(* IEC 61131-3 sources: STEPROBOT/docs/auto_job_r6_4/plc, 18 files *)

(* ---- GVL_FileBridge.st ---- *)
{attribute 'qualified_only'}
VAR_GLOBAL PERSISTENT RETAIN
    (* Reserve these MW ranges in the FIELD project before importing. *)
    aCommand AT %MW6000 : ARRAY[0..119] OF WORD;
    aHeartbeat AT %MW6120 : ARRAY[0..4] OF WORD;
    aStatus AT %MW6200 : ARRAY[0..63] OF WORD;
END_VAR
VAR_GLOBAL
    (* LOCAL configuration only. Never map credentials/permit to Modbus. *)
    xFileTransferPermit : BOOL := FALSE;
    xReset : BOOL := FALSE;
    sFtpUser : STRING(64) := '';
    sFtpPassword : STRING(64) := '';
    aBuffer : ARRAY[0..1048575] OF BYTE;
    (* One-time LOCAL commissioning: exact existing project already bound to these manual service and one auto GDI number.
       This mode reuses bindings. It never edits robot system configuration. *)
    xFixedMappingConfirmed : BOOL := FALSE;
    sFixedProject : STRING(64) := 'pcjob_manual_r63.sr';
    uiFixedCapture : UINT := UINT#10;
    uiFixedPath : UINT := UINT#11;
    uiAutoCapacity : UINT := UINT#15;
    (* Nonretained: a reboot or failed update never authorizes a partly updated project. *)
    xFixedUpdateBusy : BOOL;
    xFixedReady : BOOL;
    xFixedIdle : BOOL;
    aAutoTag : ARRAY[0..2] OF WORD;
END_VAR

(* ---- GVL_FileBridgeRetain.st ---- *)
{attribute 'qualified_only'}
VAR_GLOBAL PERSISTENT RETAIN
    udiBootCounter : UDINT := UDINT#0;
END_VAR

(* ---- GVL_ManualBridge.st ---- *)
{attribute 'qualified_only'}
VAR_GLOBAL PERSISTENT RETAIN
    // PC extension: no overlap with HR200..215, HR300..363 or FTP HR6000+.
    aCommand AT %MW220 : ARRAY[0..15] OF WORD;
    aStatus AT %MW400 : ARRAY[0..31] OF WORD;
END_VAR
VAR_GLOBAL
    // Local configuration. Assign ONE unused GDI slot to manual_service before setting TRUE.
    xInstalled : BOOL := FALSE;
    xServiceBindingConfirmed : BOOL := FALSE;
    uiServiceProgram : UINT := 10;
    // PRG_ManualBridge is the only writer. PRG_RobotBridge reads these requests.
    xActive : BOOL;
    xStartRequest : BOOL;
    xStopRequest : BOOL;
END_VAR

(* ---- GVL_ParamProbe.st ---- *)
{attribute 'qualified_only'}
VAR_GLOBAL
    // Mapped to existing ParamProbe_Write FC16 offset4 length4. Single writer: PRG_ManualBridge.
    aParamTx : ARRAY[0..3] OF WORD;
END_VAR

(* ---- GVL_RobotBridge.st ---- *)
{attribute 'qualified_only'}
VAR_GLOBAL PERSISTENT RETAIN
    // PC <-> PLC. Inovance native Modbus TCP slave: MWn <-> HR offset n.
    // Commission by reading HR300=16#4D42 and HR301=2 before permitting motion.
    aHostCmd AT %MW200 : ARRAY[0..15] OF WORD;
    aHostStatus AT %MW300 : ARRAY[0..63] OF WORD;

END_VAR

VAR_GLOBAL
    // PLC master -> STEP slave: FC04 / offset 0 / 32 WORD.
    aRobotRx : ARRAY[0..31] OF WORD;
    // PLC master -> STEP slave: ONE FC16 / offset 0 / 2 WORDs.
    // Map BOTH aRobotTx[0] and aRobotTx[1], NOT wRobotTxControl alone.
    aRobotTx : ARRAY[0..1] OF WORD;
    wRobotTxControl : WORD; // first-word diagnostic alias, not a separate channel

    // Local commissioning/operation inputs. Do not map these into aHostCmd.
    xCommissioned : BOOL := FALSE;
    // Set locally ONLY after checking DI49..56 and the GDI program bindings.
    xGdiProgramMappingConfirmed : BOOL := FALSE;
    xRemotePermit : BOOL := FALSE;
    // Optional native master/channel fault. FALSE leaves DO42 watchdog in use.
    xNativeModbusError : BOOL := FALSE;

    // Published live diagnostics.
    xRobotLinkOK : BOOL;
    xRobotRunning : BOOL;
    xRobotPaused : BOOL;
    xRobotStopped : BOOL;
    xRobotEnabled : BOOL;
    xRobotAlarm : BOOL;
    xRobotEmergency : BOOL;
    xRobotExternalAuto : BOOL;
    xHostRegistered : BOOL;
    xHostAlive : BOOL;
    xBusy : BOOL;
    xStopInterlock : BOOL;
    xLoadOperatorConfirmed : BOOL;
    uiFixedJobGuardVersion : UINT;
END_VAR

(* ---- GVL_RobotBridgeRetain.st ---- *)
{attribute 'qualified_only'}
VAR_GLOBAL PERSISTENT RETAIN
    // Incremented on application initialization, not on every scan.
    // Also require a fresh registration; a cold reset can reset RETAIN memory.
    udiBootCounter : UDINT := 0;
END_VAR

(* ---- GVL_RobotJoints.st ---- *)
{attribute 'qualified_only'}
VAR_GLOBAL PERSISTENT RETAIN
    // PC reads HR500..539. Reserve this unused range in the field project.
    // The publisher rebuilds all validity metadata; retained values never grant validity.
    aStatus AT %MW500 : ARRAY[0..39] OF WORD;
END_VAR
VAR_GLOBAL
    xEnable : BOOL := TRUE;
    sRobotAddress : STRING(15) := '192.168.3.188';
    uiRobotPort : UINT := UINT#502;
    byRobotUnit : BYTE := BYTE#1;
    // Local commissioning only: compare all six axes with the pendant.
    // FALSE = first register is the low half of IEEE754 REAL.
    xHighWordFirst : BOOL := FALSE;
END_VAR

(* ---- F_AutoFileIndex.st ---- *)
FUNCTION F_AutoFileIndex : UINT
VAR_INPUT
    sName : STRING(64);
END_VAR
F_AutoFileIndex := UINT#0;
IF sName = 'auto_main.srd' THEN F_AutoFileIndex := UINT#1; END_IF;
IF sName = 'auto_main.srp' THEN F_AutoFileIndex := UINT#2; END_IF;
IF sName = 'auto_01.srd' THEN F_AutoFileIndex := UINT#3; END_IF;
IF sName = 'auto_01.srp' THEN F_AutoFileIndex := UINT#4; END_IF;
IF sName = 'auto_02.srd' THEN F_AutoFileIndex := UINT#5; END_IF;
IF sName = 'auto_02.srp' THEN F_AutoFileIndex := UINT#6; END_IF;
IF sName = 'auto_03.srd' THEN F_AutoFileIndex := UINT#7; END_IF;
IF sName = 'auto_03.srp' THEN F_AutoFileIndex := UINT#8; END_IF;
IF sName = 'auto_04.srd' THEN F_AutoFileIndex := UINT#9; END_IF;
IF sName = 'auto_04.srp' THEN F_AutoFileIndex := UINT#10; END_IF;
IF sName = 'auto_05.srd' THEN F_AutoFileIndex := UINT#11; END_IF;
IF sName = 'auto_05.srp' THEN F_AutoFileIndex := UINT#12; END_IF;
IF sName = 'auto_06.srd' THEN F_AutoFileIndex := UINT#13; END_IF;
IF sName = 'auto_06.srp' THEN F_AutoFileIndex := UINT#14; END_IF;
IF sName = 'auto_07.srd' THEN F_AutoFileIndex := UINT#15; END_IF;
IF sName = 'auto_07.srp' THEN F_AutoFileIndex := UINT#16; END_IF;
IF sName = 'auto_08.srd' THEN F_AutoFileIndex := UINT#17; END_IF;
IF sName = 'auto_08.srp' THEN F_AutoFileIndex := UINT#18; END_IF;
IF sName = 'auto_09.srd' THEN F_AutoFileIndex := UINT#19; END_IF;
IF sName = 'auto_09.srp' THEN F_AutoFileIndex := UINT#20; END_IF;
IF sName = 'auto_10.srd' THEN F_AutoFileIndex := UINT#21; END_IF;
IF sName = 'auto_10.srp' THEN F_AutoFileIndex := UINT#22; END_IF;
IF sName = 'auto_11.srd' THEN F_AutoFileIndex := UINT#23; END_IF;
IF sName = 'auto_11.srp' THEN F_AutoFileIndex := UINT#24; END_IF;
IF sName = 'auto_12.srd' THEN F_AutoFileIndex := UINT#25; END_IF;
IF sName = 'auto_12.srp' THEN F_AutoFileIndex := UINT#26; END_IF;
IF sName = 'auto_13.srd' THEN F_AutoFileIndex := UINT#27; END_IF;
IF sName = 'auto_13.srp' THEN F_AutoFileIndex := UINT#28; END_IF;
IF sName = 'auto_14.srd' THEN F_AutoFileIndex := UINT#29; END_IF;
IF sName = 'auto_14.srp' THEN F_AutoFileIndex := UINT#30; END_IF;
IF sName = 'auto_15.srd' THEN F_AutoFileIndex := UINT#31; END_IF;
IF sName = 'auto_15.srp' THEN F_AutoFileIndex := UINT#32; END_IF;
END_FUNCTION

(* ---- F_FileCrc32.st ---- *)
FUNCTION F_FileCrc32 : UDINT
VAR_INPUT
    pData : POINTER TO BYTE;
    uiCount : UINT;
    udiSeed : UDINT;
END_VAR
VAR
    udiCrc : UDINT;
    uiI : UINT;
    uiBit : UINT;
END_VAR
(* Running reflected CRC-32. Caller supplies initial FFFFFFFF and final XOR. *)
udiCrc := udiSeed;
IF uiCount > UINT#0 THEN
    FOR uiI := UINT#0 TO uiCount - UINT#1 DO
        udiCrc := udiCrc XOR BYTE_TO_UDINT(pData[uiI]);
        FOR uiBit := UINT#0 TO UINT#7 DO
            IF (udiCrc AND UDINT#1) <> UDINT#0 THEN
                udiCrc := SHR(udiCrc, 1) XOR UDINT#16#EDB88320;
            ELSE
                udiCrc := SHR(udiCrc, 1);
            END_IF;
        END_FOR;
    END_FOR;
END_IF;
F_FileCrc32 := udiCrc;
END_FUNCTION

(* ---- F_FileCrc32Fast.st ---- *)
FUNCTION F_FileCrc32Fast : UDINT
VAR_INPUT
    pData : POINTER TO BYTE;
    uiCount : UINT;
    udiSeed : UDINT;
END_VAR
VAR
    udiCrc : UDINT;
    udiTable : UDINT;
    uiI : UINT;
    uiNibble : UINT;
END_VAR
(* Reflected CRC32, two nibble lookups per byte; no initialization scan. *)
udiCrc := udiSeed;
IF uiCount > UINT#0 THEN
    FOR uiI := UINT#0 TO uiCount - UINT#1 DO
        udiCrc := udiCrc XOR BYTE_TO_UDINT(pData[uiI]);
        FOR uiNibble := UINT#0 TO UINT#1 DO
            CASE udiCrc AND UDINT#15 OF
                0: udiTable := UDINT#16#00000000;
                1: udiTable := UDINT#16#1DB71064;
                2: udiTable := UDINT#16#3B6E20C8;
                3: udiTable := UDINT#16#26D930AC;
                4: udiTable := UDINT#16#76DC4190;
                5: udiTable := UDINT#16#6B6B51F4;
                6: udiTable := UDINT#16#4DB26158;
                7: udiTable := UDINT#16#5005713C;
                8: udiTable := UDINT#16#EDB88320;
                9: udiTable := UDINT#16#F00F9344;
                10: udiTable := UDINT#16#D6D6A3E8;
                11: udiTable := UDINT#16#CB61B38C;
                12: udiTable := UDINT#16#9B64C2B0;
                13: udiTable := UDINT#16#86D3D2D4;
                14: udiTable := UDINT#16#A00AE278;
                15: udiTable := UDINT#16#BDBDF21C;
            END_CASE;
            udiCrc := SHR(udiCrc, 4) XOR udiTable;
        END_FOR;
    END_FOR;
END_IF;
F_FileCrc32Fast := udiCrc;
END_FUNCTION

(* ---- F_FileNameValid.st ---- *)
FUNCTION F_FileNameValid : BOOL
VAR_INPUT
    sName : STRING(64);
    xProject : BOOL;
END_VAR
VAR
    pName : POINTER TO BYTE;
    uiI : UINT;
    uiBaseLength : UINT;
    xValid : BOOL;
    xChar : BOOL;
END_VAR
(* Flat lowercase ASCII names; no slash, CR/LF, spaces, or extra dots. *)
xValid := FALSE;
uiBaseLength := UINT#0;
IF xProject THEN
    IF (LEFT(sName, 6) = 'pcjob_') AND (RIGHT(sName, 3) = '.sr')
        AND (LEN(sName) >= 12) AND (LEN(sName) <= 48) THEN
        uiBaseLength := INT_TO_UINT(LEN(sName)) - UINT#3;
    END_IF;
ELSE
    IF (LEN(sName) >= 5) AND (LEN(sName) <= 48) THEN
        IF (RIGHT(sName, 4) = '.srp') OR (RIGHT(sName, 4) = '.srd')
            OR (RIGHT(sName, 4) = '.txt') THEN
            uiBaseLength := INT_TO_UINT(LEN(sName)) - UINT#4;
        END_IF;
    END_IF;
END_IF;
IF uiBaseLength > UINT#0 THEN
    xValid := TRUE;
    pName := ADR(sName);
    FOR uiI := UINT#0 TO uiBaseLength - UINT#1 DO
        xChar := ((pName[uiI] >= BYTE#97) AND (pName[uiI] <= BYTE#122))
            OR ((pName[uiI] >= BYTE#48) AND (pName[uiI] <= BYTE#57))
            OR (pName[uiI] = BYTE#95);
        IF NOT xChar THEN xValid := FALSE; END_IF;
    END_FOR;
END_IF;
F_FileNameValid := xValid;
END_FUNCTION

(* ---- F_FixedFileValid.st ---- *)
FUNCTION F_FixedFileValid : BOOL
VAR_INPUT
    sName : STRING(64);
END_VAR
F_FixedFileValid := F_AutoFileIndex(sName) > UINT#0;
END_FUNCTION

(* ---- FB_FileFtp.st ---- *)
FUNCTION_BLOCK FB_FileFtp
VAR_INPUT
    xStart : BOOL;
    xAbort : BOOL;
    pBuffer : POINTER TO BYTE;
    udiSize : UDINT;
    sProject : STRING(64);
    sFile : STRING(64);
    xCreateProject : BOOL;
    xReplaceFixed : BOOL;
    xVerifyOnly : BOOL;
    udiVerifyCrc : UDINT;
    sUser : STRING(64);
    sPassword : STRING(64);
END_VAR
VAR CONSTANT
    cdiControlID : DINT := DINT#245;
    cdiDataID : DINT := DINT#246;
END_VAR
VAR_OUTPUT
    xDone : BOOL := FALSE;
    xTestPassed : BOOL := FALSE;
    xError : BOOL := FALSE;
    xLoginOk : BOOL := FALSE;
    xBaseDirOk : BOOL := FALSE;
    xScratchCreated : BOOL := FALSE;
    xUploadComplete : BOOL := FALSE;
    xReadbackComplete : BOOL := FALSE;
    xContentMatch : BOOL := FALSE;
    xQuitOk : BOOL := FALSE;
    xCleanupOk : BOOL := FALSE;
    uiStep : UINT := UINT#0;
    uiErrorStage : UINT := UINT#0;
    wErrorID : WORD := WORD#0;
    wDataCloseErrorID : WORD := WORD#0;
    wControlCloseErrorID : WORD := WORD#0;
    udiExpectedBytes : UDINT := UDINT#0;
    udiUploadedBytes : UDINT := UDINT#0;
    udiReadbackBytes : UDINT := UDINT#0;
    uiReplyCode : UINT := UINT#0;
    uiUserReplyCode : UINT := UINT#0;
    uiPassReplyCode : UINT := UINT#0;
    uiBaseDirReplyCode : UINT := UINT#0;
    uiNameCheckReplyCode : UINT := UINT#0;
    uiMkdReplyCode : UINT := UINT#0;
    uiStorReplyCode : UINT := UINT#0;
    uiUploadCompleteCode : UINT := UINT#0;
    uiRetrReplyCode : UINT := UINT#0;
    uiDownloadCompleteCode : UINT := UINT#0;
    uiPasvPort : UINT := UINT#0;
    wReadbackEndStatus : WORD := WORD#0;
    sRemotePath : STRING(160);
    sLastReply : STRING(255);
    sMkdReply : STRING(255);
    sPasvReply : STRING(255);
    sUploadReply : STRING(255);
    sDownloadReply : STRING(255);
    xControlOwned : BOOL := FALSE;
    xDataOwned : BOOL := FALSE;
    xUploadDataConnected : BOOL := FALSE;
    xDownloadDataConnected : BOOL := FALSE;
    xLineTruncated : BOOL := FALSE;

END_VAR
VAR
    (* Caller owns immutable buffer until xDone and clean socket closure. *)
    xAbortLatched : BOOL;
    xProgress : BOOL;
    xDirectoryReady : BOOL;
    xReplaceRun : BOOL;
    sFileRun : STRING(64);
    pBufferRun : POINTER TO BYTE;

    stControlServer : CmpHCTCPIP.ADDRESS := (strIPAddr := '192.168.3.188', uiPort := UINT#21);
    stDataServer : CmpHCTCPIP.ADDRESS;
    fbControlClient : CmpHCTCPIP.SktTCPClient;
    fbControlClose : CmpHCTCPIP.SktClose;
    fbDataClient : CmpHCTCPIP.SktTCPClient;
    fbDataClose : CmpHCTCPIP.SktClose;
    fbReplyTimeout : TON;
    fbCommandTimeout : TON;
    fbUploadTimeout : TON;
    fbReadbackTimeout : TON;
    fbDataCloseTimeout : TON;
    fbControlCloseTimeout : TON;

    xStartOld : BOOL := FALSE;
    xFail : BOOL := FALSE;
    xFinishedNow : BOOL := FALSE;
    wPendingError : WORD := WORD#0;
    uiPendingStage : UINT := UINT#0;
    uiPhase : UINT := UINT#0;
    uiNextCommand : UINT := UINT#0;
    uiTransferMode : UINT := UINT#0;
    xReplyReady : BOOL := FALSE;
    xReplyAccepted : BOOL := FALSE;
    xDigits : BOOL := FALSE;
    xMultiline : BOOL := FALSE;
    sMultilineCode : STRING(3);
    sLine : STRING(255);
    pLine : POINTER TO BYTE;
    uiLineLength : UINT := UINT#0;
    fbControlIo : FB_FileSocketIo;
    fbDataIo : FB_FileSocketIo;
    uiControlRxIndex : UINT;
    uiControlRxCount : UINT;
    uiParse : UINT;
    byControl : BYTE;
    pSendNow : POINTER TO BYTE;
    uiSendNow : UINT;
    xVerifyRun : BOOL;
    udiVerifyCrcRun : UDINT;
    udiReadbackCrc : UDINT;
    sCommand : STRING(160);
    pCommand : POINTER TO BYTE;
    uiCommandIndex : UINT := UINT#0;
    uiCommandLength : UINT := UINT#0;
    sUserRun : STRING(64);
    sPasswordRun : STRING(64);
    sScratchRun : STRING(64);
    pCredential : POINTER TO BYTE;
    uiI : UINT := UINT#0;
    xNameCharacter : BOOL := FALSE;
    xBytesMatch : BOOL := FALSE;
    xReadbackEndCandidate : BOOL := FALSE;
    xDataCloseFailed : BOOL := FALSE;
    pReply : POINTER TO BYTE;
    aPasv : ARRAY[0..5] OF UINT;
    uiPasvField : UINT := UINT#0;
    uiPasvValue : UINT := UINT#0;
    xPasvValid : BOOL := FALSE;
    xPasvInTuple : BOOL := FALSE;
    xPasvClosed : BOOL := FALSE;
    xPasvHasDigit : BOOL := FALSE;
END_VAR
(* Derived from field-passed PRG_FtpUploadProbe. New bridge is NOT field validated. *)
(* IDs 245/246 must be free; default cabinet 192.168.3.188:21. *)
(* Bounded 8192-byte I/O, exact offsets and explicit EOF. No motion commands. *)
pLine := ADR(sLine);
pCommand := ADR(sCommand);
xFail := FALSE;
xFinishedNow := FALSE;
xReplyReady := FALSE;
wPendingError := WORD#0;
uiPendingStage := UINT#20 + uiPhase * UINT#10;

pSendNow := pCommand;
uiSendNow := UINT#0;
IF uiStep = UINT#40 THEN
    pSendNow := pCommand + uiCommandIndex;
    uiSendNow := uiCommandLength - uiCommandIndex;
END_IF;
fbControlClient(xExecute := uiStep = UINT#10, diConnectID := cdiControlID,
    stServerAddress := stControlServer);
fbControlIo(xSend := uiStep = UINT#40,
    xReceive := (uiStep = UINT#20) AND (uiControlRxIndex >= uiControlRxCount),
    diConnectID := cdiControlID, pSend := pSendNow, uiSendSize := uiSendNow);
IF fbControlIo.uiCount > UINT#0 THEN
    uiControlRxIndex := UINT#0;
    uiControlRxCount := fbControlIo.uiCount;
END_IF;
pSendNow := pBufferRun;
uiSendNow := UINT#0;
IF (uiStep = UINT#60) AND (udiUploadedBytes < udiExpectedBytes) THEN
    pSendNow := pBufferRun + udiUploadedBytes;
    IF udiExpectedBytes - udiUploadedBytes > UDINT#8192 THEN
        uiSendNow := UINT#8192;
    ELSE
        uiSendNow := UDINT_TO_UINT(udiExpectedBytes - udiUploadedBytes);
    END_IF;
END_IF;
fbDataClient(xExecute := uiStep = UINT#50, diConnectID := cdiDataID,
    stServerAddress := stDataServer);
fbDataIo(xSend := (uiStep = UINT#60) AND (uiSendNow > UINT#0),
    xReceive := uiStep = UINT#70, diConnectID := cdiDataID,
    pSend := pSendNow, uiSendSize := uiSendNow);
fbDataClose(xExecute := ((uiStep = UINT#80) OR (uiStep = UINT#90))
    AND xDataOwned AND NOT xDataCloseFailed, diConnectID := cdiDataID);
fbControlClose(xExecute := (uiStep = UINT#95) AND xControlOwned,
    diConnectID := cdiControlID);
fbReplyTimeout(IN := uiStep = UINT#20, PT := T#20s);
fbCommandTimeout(IN := (uiStep = UINT#40) OR (uiStep = UINT#45), PT := T#30s);
xProgress := ((uiStep = UINT#60) AND (fbDataIo.uiSent > UINT#0))
    OR ((uiStep = UINT#70) AND (fbDataIo.uiCount > UINT#0));
fbUploadTimeout(IN := ((uiStep = UINT#60) OR (uiStep = UINT#65)) AND NOT xProgress,
    PT := T#30s);
fbReadbackTimeout(IN := (uiStep = UINT#70) AND NOT xProgress, PT := T#30s);
fbDataCloseTimeout(IN := ((uiStep = UINT#80) OR (uiStep = UINT#90))
    AND xDataOwned AND NOT xDataCloseFailed, PT := T#5s);
fbControlCloseTimeout(IN := uiStep = UINT#95, PT := T#5s);

(* Bounded control-reply parser; identical-code SPACE terminates multiline replies. *)
IF (uiStep = UINT#20) AND NOT fbControlIo.xError THEN
    IF uiControlRxIndex < uiControlRxCount THEN
    FOR uiParse := uiControlRxIndex TO uiControlRxCount - UINT#1 DO
      IF (uiControlRxIndex < uiControlRxCount) AND NOT xReplyReady AND NOT xFail THEN
        byControl := fbControlIo.aRecv[uiControlRxIndex];
        uiControlRxIndex := uiControlRxIndex + UINT#1;
        IF byControl = BYTE#10 THEN
            IF uiLineLength > UINT#0 THEN
                IF pLine[uiLineLength - UINT#1] = BYTE#13 THEN
                    uiLineLength := uiLineLength - UINT#1;
                    pLine[uiLineLength] := BYTE#0;
                END_IF;
            END_IF;
            IF xMultiline THEN
                IF LEFT(sLine, 4) = CONCAT(sMultilineCode, ' ') THEN
                    xMultiline := FALSE;
                    xReplyReady := TRUE;
                END_IF;
            ELSE
                xDigits := FALSE;
                IF uiLineLength >= UINT#4 THEN
                    xDigits := (pLine[0] >= BYTE#48) AND (pLine[0] <= BYTE#57)
                        AND (pLine[1] >= BYTE#48) AND (pLine[1] <= BYTE#57)
                        AND (pLine[2] >= BYTE#48) AND (pLine[2] <= BYTE#57);
                END_IF;
                IF xDigits THEN
                    IF pLine[3] = BYTE#45 THEN
                        xMultiline := TRUE;
                        sMultilineCode := LEFT(sLine, 3);
                    ELSIF pLine[3] = BYTE#32 THEN
                        xReplyReady := TRUE;
                    ELSE
                        xFail := TRUE;
                        wPendingError := WORD#16#F203;
                    END_IF;
                ELSE
                    xFail := TRUE;
                    wPendingError := WORD#16#F203;
                END_IF;
            END_IF;
            IF xReplyReady THEN
                uiReplyCode := (BYTE_TO_UINT(pLine[0]) - UINT#48) * UINT#100
                    + (BYTE_TO_UINT(pLine[1]) - UINT#48) * UINT#10
                    + BYTE_TO_UINT(pLine[2]) - UINT#48;
                sLastReply := sLine;
            ELSIF xFail THEN
                sLastReply := sLine;
            END_IF;
            sLine := '';
            uiLineLength := UINT#0;
        ELSE
            IF uiLineLength < UINT#255 THEN
                pLine[uiLineLength] := byControl;
                uiLineLength := uiLineLength + UINT#1;
                pLine[uiLineLength] := BYTE#0;
            ELSE
                xLineTruncated := TRUE;
                sLastReply := sLine;
                xFail := TRUE;
                wPendingError := WORD#16#F204;
            END_IF;
        END_IF;
      END_IF;
    END_FOR;
    END_IF;
END_IF;

CASE uiStep OF
    UINT#0:
        IF xStart AND NOT xStartOld THEN
            xAbortLatched := FALSE;
            xDirectoryReady := FALSE;
            xDone := FALSE;
            xTestPassed := FALSE;
            xError := FALSE;
            xLoginOk := FALSE;
            xBaseDirOk := FALSE;
            xScratchCreated := FALSE;
            xUploadComplete := FALSE;
            xReadbackComplete := FALSE;
            xContentMatch := FALSE;
            xQuitOk := FALSE;
            xCleanupOk := FALSE;
            xUploadDataConnected := FALSE;
            xDownloadDataConnected := FALSE;
            xDataCloseFailed := FALSE;
            xLineTruncated := FALSE;
            xReadbackEndCandidate := FALSE;
            xBytesMatch := TRUE;
            uiErrorStage := UINT#0;
            wErrorID := WORD#0;
            wDataCloseErrorID := WORD#0;
            wControlCloseErrorID := WORD#0;
            wReadbackEndStatus := WORD#0;
            udiUploadedBytes := UDINT#0;
            udiReadbackBytes := UDINT#0;
            uiReplyCode := UINT#0;
            uiUserReplyCode := UINT#0;
            uiPassReplyCode := UINT#0;
            uiBaseDirReplyCode := UINT#0;
            uiNameCheckReplyCode := UINT#0;
            uiMkdReplyCode := UINT#0;
            uiStorReplyCode := UINT#0;
            uiUploadCompleteCode := UINT#0;
            uiRetrReplyCode := UINT#0;
            uiDownloadCompleteCode := UINT#0;
            uiPasvPort := UINT#0;
            sLastReply := '';
            sMkdReply := '';
            sPasvReply := '';
            sUploadReply := '';
            sDownloadReply := '';
            sLine := '';
            uiLineLength := UINT#0;
            uiControlRxIndex := UINT#0;
            uiControlRxCount := UINT#0;
            xMultiline := FALSE;
            sMultilineCode := '';
            uiPhase := UINT#0;
            uiTransferMode := UINT#0;
            sUserRun := sUser;
            sPasswordRun := sPassword;
            sScratchRun := sProject;
            sFileRun := sFile;
            xReplaceRun := xReplaceFixed;
            xVerifyRun := xVerifyOnly;
            udiVerifyCrcRun := udiVerifyCrc;
            udiReadbackCrc := UDINT#16#FFFFFFFF;
            pBufferRun := pBuffer;
            sRemotePath := CONCAT(CONCAT(CONCAT('/UserPrograms/', sScratchRun), '/'), sFileRun);
            udiExpectedBytes := udiSize;
            uiPendingStage := UINT#1;
            IF (LEN(sUserRun) = 0) OR (LEN(sPasswordRun) = 0) THEN
                xFail := TRUE;
                wPendingError := WORD#16#F200;
            ELSE
                pCredential := ADR(sUserRun);
                FOR uiI := UINT#0 TO INT_TO_UINT(LEN(sUserRun)) - UINT#1 DO
                    IF (pCredential[uiI] < BYTE#32) OR (pCredential[uiI] > BYTE#126) THEN
                        xFail := TRUE;
                        wPendingError := WORD#16#F207;
                    END_IF;
                END_FOR;
                pCredential := ADR(sPasswordRun);
                FOR uiI := UINT#0 TO INT_TO_UINT(LEN(sPasswordRun)) - UINT#1 DO
                    IF (pCredential[uiI] < BYTE#32) OR (pCredential[uiI] > BYTE#126) THEN
                        xFail := TRUE;
                        wPendingError := WORD#16#F207;
                    END_IF;
                END_FOR;
            END_IF;
            IF NOT F_FileNameValid(sScratchRun, TRUE)
                OR NOT F_FileNameValid(sFileRun, FALSE)
                OR (udiExpectedBytes > UDINT#1048576)
                OR (pBufferRun = 0) THEN
                xFail := TRUE;
                wPendingError := WORD#16#F209;
            END_IF;
            IF xVerifyRun AND NOT xReplaceRun THEN
                xFail := TRUE;
                wPendingError := WORD#16#F20C;
            END_IF;
            IF xReplaceRun AND (NOT GVL_FileBridge.xFixedMappingConfirmed
                OR (GVL_RobotBridge.uiFixedJobGuardVersion <> UINT#140)
                OR NOT GVL_FileBridge.xFixedIdle OR (sScratchRun <> GVL_FileBridge.sFixedProject)
                OR NOT F_FixedFileValid(sFileRun)) THEN
                xFail := TRUE;
                wPendingError := WORD#16#F20C;
            END_IF;
            IF NOT xFail THEN
                uiStep := UINT#10;
            END_IF;
        END_IF;

    UINT#10:
        IF fbControlClient.xError THEN
            xFail := TRUE;
            wPendingError := fbControlClient.wErrorID;
            uiPendingStage := UINT#10;
        ELSIF fbControlClient.xDone THEN
            xControlOwned := TRUE;
            uiStep := UINT#20;
        END_IF;

    UINT#20:
        IF fbControlIo.xError OR fbControlIo.xPeerClosed THEN
            xFail := TRUE;
            wPendingError := WORD#16#F224;
        ELSIF NOT xFail THEN
            IF xReplyReady THEN
                xReplyAccepted := FALSE;
                CASE uiPhase OF
                    UINT#0:
                        IF uiReplyCode = UINT#220 THEN
                            xReplyAccepted := TRUE;
                            uiNextCommand := UINT#1;
                            uiStep := UINT#30;
                        ELSIF uiReplyCode = UINT#140 THEN
                            xReplyAccepted := TRUE;
                        END_IF;
                    UINT#1:
                        uiUserReplyCode := uiReplyCode;
                        IF uiReplyCode = UINT#331 THEN
                            xReplyAccepted := TRUE;
                            uiNextCommand := UINT#2;
                            uiStep := UINT#30;
                        ELSIF uiReplyCode = UINT#230 THEN
                            xReplyAccepted := TRUE;
                            xLoginOk := TRUE;
                            uiNextCommand := UINT#3;
                            uiStep := UINT#30;
                        END_IF;
                    UINT#2:
                        uiPassReplyCode := uiReplyCode;
                        IF uiReplyCode = UINT#230 THEN
                            xReplyAccepted := TRUE;
                            xLoginOk := TRUE;
                            uiNextCommand := UINT#3;
                            uiStep := UINT#30;
                        END_IF;
                    UINT#3:
                        uiBaseDirReplyCode := uiReplyCode;
                        IF uiReplyCode = UINT#250 THEN
                            xReplyAccepted := TRUE;
                            xBaseDirOk := TRUE;
                            IF xCreateProject OR xReplaceRun THEN
                                uiNextCommand := UINT#14;
                            ELSE
                                uiNextCommand := UINT#5;
                            END_IF;
                            uiStep := UINT#30;
                        END_IF;
                    UINT#14:
                        uiNameCheckReplyCode := uiReplyCode;
                        IF uiReplyCode = UINT#550 THEN
                            xReplyAccepted := TRUE;
                            IF xReplaceRun THEN
                                (* Fixed binding must already exist: never silently create another target. *)
                                xFail := TRUE;
                                wPendingError := WORD#16#F20B;
                            ELSE
                                uiNextCommand := UINT#4;
                                uiStep := UINT#30;
                            END_IF;
                        ELSIF uiReplyCode = UINT#250 THEN
                            xReplyAccepted := TRUE;
                            IF xReplaceRun THEN
                                xDirectoryReady := TRUE;
                                uiNextCommand := UINT#6;
                                uiStep := UINT#30;
                            ELSE
                                (* Original mode retains its no-overwrite behavior. *)
                                xFail := TRUE;
                                wPendingError := WORD#16#F208;
                            END_IF;
                        END_IF;
                    UINT#4:
                        uiMkdReplyCode := uiReplyCode;
                        sMkdReply := sLastReply;
                        IF uiReplyCode = UINT#257 THEN
                            xReplyAccepted := TRUE;
                            xScratchCreated := TRUE;
                            uiNextCommand := UINT#5;
                            uiStep := UINT#30;
                        END_IF;
                    UINT#5:
                        IF uiReplyCode = UINT#250 THEN
                            xDirectoryReady := TRUE;
                            xReplyAccepted := TRUE;
                            uiNextCommand := UINT#6;
                            uiStep := UINT#30;
                        END_IF;
                    UINT#6:
                        IF uiReplyCode = UINT#200 THEN
                            xReplyAccepted := TRUE;
                            IF xVerifyRun THEN uiNextCommand := UINT#10;
                            ELSE uiNextCommand := UINT#7; END_IF;
                            uiStep := UINT#30;
                        END_IF;
                    UINT#7, UINT#10:
                        IF uiReplyCode = UINT#227 THEN
                            xReplyAccepted := TRUE;
                            sPasvReply := sLastReply;
                            uiStep := UINT#35;
                        END_IF;
                    UINT#8:
                        uiStorReplyCode := uiReplyCode;
                        IF (uiReplyCode = UINT#125) OR (uiReplyCode = UINT#150) THEN
                            xReplyAccepted := TRUE;
                            IF udiExpectedBytes = UDINT#0 THEN
                                (* Empty STOR still needs data EOF, 226 and exact RETR. *)
                                uiStep := UINT#80;
                            ELSE
                                uiStep := UINT#60;
                            END_IF;
                        END_IF;
                    UINT#9:
                        uiUploadCompleteCode := uiReplyCode;
                        sUploadReply := sLastReply;
                        IF (uiReplyCode = UINT#226) OR (uiReplyCode = UINT#250) THEN
                            xReplyAccepted := TRUE;
                            xUploadComplete := TRUE;
                            uiNextCommand := UINT#10;
                            uiStep := UINT#30;
                        END_IF;
                    UINT#11:
                        uiRetrReplyCode := uiReplyCode;
                        IF (uiReplyCode = UINT#125) OR (uiReplyCode = UINT#150) THEN
                            xReplyAccepted := TRUE;
                            uiStep := UINT#70;
                        END_IF;
                    UINT#12:
                        uiDownloadCompleteCode := uiReplyCode;
                        sDownloadReply := sLastReply;
                        IF (uiReplyCode = UINT#226) OR (uiReplyCode = UINT#250) THEN
                            xReplyAccepted := TRUE;
                            xReadbackComplete := TRUE;
                            xContentMatch := xBytesMatch AND xReadbackEndCandidate
                                AND (udiReadbackBytes = udiExpectedBytes);
                            IF xContentMatch THEN
                                uiNextCommand := UINT#13;
                                uiStep := UINT#30;
                            ELSE
                                xFail := TRUE;
                                wPendingError := WORD#16#F205;
                            END_IF;
                        END_IF;
                    UINT#13:
                        IF uiReplyCode = UINT#221 THEN
                            xReplyAccepted := TRUE;
                            xQuitOk := TRUE;
                            uiStep := UINT#90;
                        END_IF;
                END_CASE;
                IF NOT xReplyAccepted THEN
                    xFail := TRUE;
                    wPendingError := WORD#16#F202;
                END_IF;
            ELSIF fbReplyTimeout.Q THEN
                xFail := TRUE;
                wPendingError := WORD#16#F201;
            END_IF;
        END_IF;

    UINT#30:
        uiPhase := uiNextCommand;
        CASE uiNextCommand OF
            UINT#1: sCommand := CONCAT(CONCAT('USER ', sUserRun), '$R$N');
            UINT#2: sCommand := CONCAT(CONCAT('PASS ', sPasswordRun), '$R$N');
            UINT#3: sCommand := 'CWD /UserPrograms$R$N';
            UINT#4: sCommand := CONCAT(CONCAT('MKD ', sScratchRun), '$R$N');
            UINT#5, UINT#14: sCommand := CONCAT(CONCAT('CWD ', sScratchRun), '$R$N');
            UINT#6: sCommand := 'TYPE I$R$N';
            UINT#7, UINT#10: sCommand := 'PASV$R$N';
            UINT#8: sCommand := CONCAT(CONCAT('STOR ', sFileRun), '$R$N');
            UINT#11: sCommand := CONCAT(CONCAT('RETR ', sFileRun), '$R$N');
            UINT#13: sCommand := 'QUIT$R$N';
        ELSE
            xFail := TRUE;
            wPendingError := WORD#16#F20A;
        END_CASE;
        IF NOT xFail THEN
            uiCommandLength := INT_TO_UINT(LEN(sCommand));
            uiCommandIndex := UINT#0;
            uiStep := UINT#40;
        END_IF;

    UINT#35:
        (* Parse six decimal octets in the first parenthesized PASV tuple. *)
        pReply := ADR(sPasvReply);
        xPasvValid := TRUE;
        xPasvInTuple := FALSE;
        xPasvClosed := FALSE;
        xPasvHasDigit := FALSE;
        uiPasvField := UINT#0;
        uiPasvValue := UINT#0;
        FOR uiI := UINT#0 TO INT_TO_UINT(LEN(sPasvReply)) - UINT#1 DO
            IF NOT xPasvInTuple THEN
                IF pReply[uiI] = BYTE#40 THEN
                    xPasvInTuple := TRUE;
                END_IF;
            ELSIF NOT xPasvClosed THEN
                IF (pReply[uiI] >= BYTE#48) AND (pReply[uiI] <= BYTE#57) THEN
                    xPasvHasDigit := TRUE;
                    IF uiPasvValue <= UINT#255 THEN
                        uiPasvValue := uiPasvValue * UINT#10 + BYTE_TO_UINT(pReply[uiI]) - UINT#48;
                        IF uiPasvValue > UINT#255 THEN
                            xPasvValid := FALSE;
                        END_IF;
                    ELSE
                        xPasvValid := FALSE;
                    END_IF;
                ELSIF (pReply[uiI] = BYTE#44) OR (pReply[uiI] = BYTE#41) THEN
                    IF NOT xPasvHasDigit OR (uiPasvField > UINT#5) OR (uiPasvValue > UINT#255) THEN
                        xPasvValid := FALSE;
                    ELSE
                        aPasv[uiPasvField] := uiPasvValue;
                        uiPasvField := uiPasvField + UINT#1;
                    END_IF;
                    uiPasvValue := UINT#0;
                    xPasvHasDigit := FALSE;
                    IF pReply[uiI] = BYTE#41 THEN
                        xPasvClosed := TRUE;
                    END_IF;
                ELSE
                    xPasvValid := FALSE;
                END_IF;
            END_IF;
        END_FOR;
        IF NOT xPasvInTuple OR NOT xPasvClosed OR (uiPasvField <> UINT#6) THEN
            xPasvValid := FALSE;
        END_IF;
        IF xPasvValid THEN
            uiPasvPort := aPasv[4] * UINT#256 + aPasv[5];
            IF (uiPasvPort = UINT#0) OR (uiPasvPort = UINT#21) THEN
                xPasvValid := FALSE;
            END_IF;
        END_IF;
        IF xPasvValid THEN
            (* Data connections are pinned to the control server, not a third-party PASV IP. *)
            stDataServer.strIPAddr := stControlServer.strIPAddr;
            stDataServer.uiPort := uiPasvPort;
            xDataCloseFailed := FALSE;
            IF uiPhase = UINT#7 THEN
                uiTransferMode := UINT#1;
            ELSE
                uiTransferMode := UINT#2;
            END_IF;
            uiStep := UINT#50;
        ELSE
            xFail := TRUE;
            wPendingError := WORD#16#F20B;
        END_IF;

    UINT#40:
        IF fbControlIo.xError THEN
            xFail := TRUE;
            wPendingError := fbControlIo.wErrorID;
        ELSIF fbControlIo.uiSent > UINT#0 THEN
            uiCommandIndex := uiCommandIndex + fbControlIo.uiSent;
            IF uiCommandIndex = uiCommandLength THEN
                sCommand := '';
                uiStep := UINT#20;
            END_IF;
        ELSIF fbCommandTimeout.Q THEN
            xFail := TRUE;
            wPendingError := WORD#16#F206;
        END_IF;

    UINT#50:
        uiPendingStage := UINT#200 + uiTransferMode;
        IF fbDataClient.xError THEN
            xFail := TRUE;
            wPendingError := fbDataClient.wErrorID;
        ELSIF fbDataClient.xDone THEN
            xDataOwned := TRUE;
            IF uiTransferMode = UINT#1 THEN
                xUploadDataConnected := TRUE;
                uiNextCommand := UINT#8;
            ELSE
                xDownloadDataConnected := TRUE;
                uiNextCommand := UINT#11;
            END_IF;
            uiStep := UINT#30;
        END_IF;

    UINT#60:
        uiPendingStage := UINT#210;
        IF fbDataIo.xError THEN
            xFail := TRUE;
            wPendingError := fbDataIo.wErrorID;
        ELSIF fbDataIo.uiSent > UINT#0 THEN
            udiUploadedBytes := udiUploadedBytes + UINT_TO_UDINT(fbDataIo.uiSent);
            IF udiUploadedBytes = udiExpectedBytes THEN uiStep := UINT#80; END_IF;
        ELSIF fbUploadTimeout.Q THEN
            xFail := TRUE;
            wPendingError := WORD#16#F206;
        END_IF;

    UINT#70:
        uiPendingStage := UINT#220;
        IF fbDataIo.xError THEN
            xFail := TRUE;
            wPendingError := fbDataIo.wErrorID;
        ELSIF fbDataIo.uiCount > UINT#0 THEN
            IF UINT_TO_UDINT(fbDataIo.uiCount) > udiExpectedBytes - udiReadbackBytes THEN
                xBytesMatch := FALSE;
                xFail := TRUE;
                wPendingError := WORD#16#F205;
            ELSE
                IF xVerifyRun THEN
                    udiReadbackCrc := F_FileCrc32Fast(ADR(fbDataIo.aRecv), fbDataIo.uiCount, udiReadbackCrc);
                ELSE
                    FOR uiI := UINT#0 TO fbDataIo.uiCount - UINT#1 DO
                        IF fbDataIo.aRecv[uiI] <> pBufferRun[udiReadbackBytes + UINT_TO_UDINT(uiI)] THEN
                            xBytesMatch := FALSE;
                        END_IF;
                    END_FOR;
                END_IF;
                udiReadbackBytes := udiReadbackBytes + UINT_TO_UDINT(fbDataIo.uiCount);
                IF NOT xBytesMatch THEN
                    xFail := TRUE;
                    wPendingError := WORD#16#F205;
                END_IF;
            END_IF;
        ELSIF fbDataIo.xPeerClosed THEN
            IF xVerifyRun AND ((udiReadbackCrc XOR UDINT#16#FFFFFFFF) <> udiVerifyCrcRun) THEN
                xBytesMatch := FALSE;
            END_IF;
            IF xBytesMatch AND (udiReadbackBytes = udiExpectedBytes) THEN
                xReadbackEndCandidate := TRUE;
                uiStep := UINT#80;
            ELSE
                xFail := TRUE;
                wPendingError := WORD#16#F205;
            END_IF;
        ELSIF fbReadbackTimeout.Q THEN
            xFail := TRUE;
            wPendingError := WORD#16#F201;
        END_IF;

    UINT#80:
        IF fbDataClose.xError OR fbDataCloseTimeout.Q THEN
            IF fbDataClose.xError THEN
                wDataCloseErrorID := fbDataClose.wErrorID;
            ELSE
                wDataCloseErrorID := WORD#16#F20C;
            END_IF;
            xDataCloseFailed := TRUE;
            IF NOT xError THEN
                xError := TRUE;
                wErrorID := wDataCloseErrorID;
                uiErrorStage := UINT#290;
            END_IF;
            uiStep := UINT#95;
        ELSIF fbDataClose.xDone THEN
            xDataOwned := FALSE;
            IF uiTransferMode = UINT#1 THEN
                uiPhase := UINT#9;
            ELSE
                uiPhase := UINT#12;
            END_IF;
            uiStep := UINT#20;
        END_IF;

    UINT#90:
        IF NOT xDataOwned OR xDataCloseFailed THEN
            uiStep := UINT#95;
        ELSIF fbDataClose.xError OR fbDataCloseTimeout.Q THEN
            IF fbDataClose.xError THEN
                wDataCloseErrorID := fbDataClose.wErrorID;
            ELSE
                wDataCloseErrorID := WORD#16#F20C;
            END_IF;
            xDataCloseFailed := TRUE;
            IF NOT xError THEN
                xError := TRUE;
                wErrorID := wDataCloseErrorID;
                uiErrorStage := UINT#290;
            END_IF;
            uiStep := UINT#95;
        ELSIF fbDataClose.xDone THEN
            xDataOwned := FALSE;
            uiStep := UINT#95;
        END_IF;

    UINT#95:
        IF NOT xControlOwned THEN
            xDone := TRUE;
            xFinishedNow := TRUE;
            uiStep := UINT#100;
        ELSIF fbControlClose.xError OR fbControlCloseTimeout.Q THEN
            IF fbControlClose.xError THEN
                wControlCloseErrorID := fbControlClose.wErrorID;
            ELSE
                wControlCloseErrorID := WORD#16#F20C;
            END_IF;
            IF NOT xError THEN
                xError := TRUE;
                wErrorID := wControlCloseErrorID;
                uiErrorStage := UINT#295;
            END_IF;
            xDone := TRUE;
            xFinishedNow := TRUE;
            uiStep := UINT#100;
        ELSIF fbControlClose.xDone THEN
            xControlOwned := FALSE;
            xDone := TRUE;
            xFinishedNow := TRUE;
            uiStep := UINT#100;
        END_IF;

    UINT#100:
        IF NOT xStart AND NOT xControlOwned AND NOT xDataOwned THEN
            uiStep := UINT#0;
        END_IF;
END_CASE;

(* Never cancel a pending native connect before its terminal result. *)
IF xAbort AND (uiStep <> UINT#0) AND (uiStep <> UINT#100) THEN
    xAbortLatched := TRUE;
END_IF;
IF xAbortLatched AND (uiStep <> UINT#0) AND (uiStep <> UINT#10)
    AND (uiStep <> UINT#50) AND (uiStep <> UINT#90)
    AND (uiStep <> UINT#95) AND (uiStep <> UINT#100) THEN
    xFail := TRUE;
    wPendingError := WORD#16#F20D;
END_IF;
IF xFail THEN
    IF NOT xError THEN
        xError := TRUE;
        wErrorID := wPendingError;
        uiErrorStage := uiPendingStage;
    END_IF;
    uiStep := UINT#90;
END_IF;

IF xFinishedNow THEN
    xCleanupOk := NOT xControlOwned AND NOT xDataOwned
        AND (wDataCloseErrorID = WORD#0) AND (wControlCloseErrorID = WORD#0);
    xTestPassed := xLoginOk AND xBaseDirOk AND xDirectoryReady
        AND (xVerifyRun OR xUploadDataConnected) AND xDownloadDataConnected
        AND (xVerifyRun OR xUploadComplete) AND xReadbackComplete AND xContentMatch
        AND xQuitOk AND xCleanupOk AND NOT xError;
    sPasswordRun := '';
    sUserRun := '';
    sCommand := '';
END_IF;
xStartOld := xStart;
END_FUNCTION_BLOCK

(* ---- FB_FileSocketIo.st ---- *)
FUNCTION_BLOCK FB_FileSocketIo
VAR_INPUT
    xSend : BOOL;
    xReceive : BOOL;
    diConnectID : DINT;
    pSend : POINTER TO BYTE;
    uiSendSize : UINT;
END_VAR
VAR_OUTPUT
    uiSent : UINT;
    uiCount : UINT;
    xPeerClosed : BOOL;
    xError : BOOL;
    wErrorID : WORD;
    udiNativeResult : UDINT;
    aRecv : ARRAY[0..8191] OF BYTE;
END_VAR
VAR
    stSocketInfo : CmpHCTCPIP.SOCKET_INFO;
    wLookup : WORD;
    xiCount : __XINT;
END_VAR
(* CmpHCTCPIP 1.0.0.7 owns the connection. This block only performs I/O.
   One nonblocking syscall per call. Parent advances by the ACTUAL count.
   No reset scan; no re-send of an already accepted prefix; EOF is explicit. *)
uiSent := UINT#0;
uiCount := UINT#0;
xPeerClosed := FALSE;
xError := FALSE;
wErrorID := WORD#0;
(* Preserve the last native result/count while idle for field diagnostics. *)
IF xSend OR xReceive THEN
    udiNativeResult := UDINT#0;
    wLookup := CmpHCTCPIP.GetSocketInfo(diConnectID, ADR(stSocketInfo));
    IF wLookup <> WORD#0 THEN
        xError := TRUE;
        wErrorID := wLookup;
    ELSIF (stSocketInfo.hSocket = SysSocket.RTS_INVALID_HANDLE)
        OR (stSocketInfo.diSocketType <> SysSocket.SOCKET_STREAM) OR (xSend AND xReceive) THEN
        xError := TRUE;
        wErrorID := WORD#16#F220;
    ELSIF xSend THEN
        IF (pSend = 0) OR (uiSendSize = UINT#0) OR (uiSendSize > UINT#8192) THEN
            xError := TRUE;
            wErrorID := WORD#16#F221;
        ELSE
            xiCount := SysSocket.SysSockSend(stSocketInfo.hSocket, pSend,
                UINT_TO_DINT(uiSendSize), SysSocket.SOCKET_MSG_DONTWAIT, ADR(udiNativeResult));
            IF udiNativeResult = CmpErrors.Errors.ERR_SOCK_WOULDBLOCK THEN
                (* Retry on the next PLC scan; the parent enforces the progress timeout. *)
            ELSIF (udiNativeResult <> CmpErrors.Errors.ERR_OK) OR (xiCount <= 0)
                OR (xiCount > UINT_TO_DINT(uiSendSize)) THEN
                xError := TRUE;
                wErrorID := WORD#16#F222;
            ELSE
                uiSent := __XINT_TO_UINT(xiCount);
            END_IF;
        END_IF;
    ELSE
        xiCount := SysSocket.SysSockRecv(stSocketInfo.hSocket, ADR(aRecv),
            DINT#8192, SysSocket.SOCKET_MSG_DONTWAIT, ADR(udiNativeResult));
        IF udiNativeResult = CmpErrors.Errors.ERR_SOCK_WOULDBLOCK THEN
            (* No data yet. A short final packet is delivered immediately. *)
        ELSIF (udiNativeResult = CmpErrors.Errors.ERR_SOCK_CLOSED) AND (xiCount = 0) THEN
            (* CODESYS reports a graceful TCP end with ERR_SOCK_CLOSED.
               Parent still requires exact length/content, FTP 226/250 and cleanup. *)
            xPeerClosed := TRUE;
        ELSIF (udiNativeResult <> CmpErrors.Errors.ERR_OK) OR (xiCount < 0) OR (xiCount > 8192) THEN
            xError := TRUE;
            wErrorID := WORD#16#F223;
        ELSIF xiCount = 0 THEN
            xPeerClosed := TRUE;
        ELSE
            uiCount := __XINT_TO_UINT(xiCount);
        END_IF;
    END_IF;
END_IF;
END_FUNCTION_BLOCK

(* ---- FB_RobotJointRead.st ---- *)
FUNCTION_BLOCK FB_RobotJointRead
VAR_INPUT
    xEnable : BOOL;
    sAddress : STRING(15);
    uiPort : UINT;
    byUnit : BYTE;
END_VAR
VAR_OUTPUT
    xValid : BOOL;
    xError : BOOL;
    xCleanupFault : BOOL;
    wErrorID : WORD;
    uiStep : UINT;
    udiCounter : UDINT;
    uiAgeMs : UINT;
    aWords : ARRAY[0..11] OF WORD;
END_VAR
VAR CONSTANT
    // Dedicated read-only socket. Never share with FTP IDs245/246.
    cdiConnectID : DINT := DINT#244;
END_VAR
VAR
    stServer : CmpHCTCPIP.ADDRESS;
    fbClient : CmpHCTCPIP.SktTCPClient;
    fbClose : CmpHCTCPIP.SktClose;
    fbIo : FB_FileSocketIo;
    fbReplyTime : TON;
    fbCloseTime : TON;
    fbPollTime : TON;
    fbRetryTime : TON;
    fbAge : TON;
    xOwned : BOOL;
    xStop : BOOL;
    xUpdated : BOOL;
    xFail : BOOL;
    sRunAddress : STRING(15);
    uiRunPort : UINT;
    byRunUnit : BYTE;
    uiTransaction : UINT;
    uiSent : UINT;
    uiReceived : UINT;
    uiSendSize : UINT;
    pSend : POINTER TO BYTE;
    aRequest : ARRAY[0..11] OF BYTE;
    aResponse : ARRAY[0..32] OF BYTE;
    i : UINT;
END_VAR
// A persistent TCP connection performs ONLY FC04 / offset64 / count12.
// No registration, parameters, program loading, enable or motion commands.
xUpdated := FALSE;
xFail := FALSE;
xStop := NOT xEnable OR (sAddress <> sRunAddress)
    OR (uiPort <> uiRunPort) OR (byUnit <> byRunUnit);
IF xStop THEN xValid := FALSE; END_IF;
pSend := ADR(aRequest);
uiSendSize := UINT#0;
IF uiStep = UINT#30 THEN
    pSend := ADR(aRequest) + uiSent;
    uiSendSize := UINT#12 - uiSent;
END_IF;
fbClient(xExecute := uiStep = UINT#10, diConnectID := cdiConnectID,
    stServerAddress := stServer);
fbIo(xSend := (uiStep = UINT#30) AND NOT xStop,
    xReceive := (uiStep = UINT#40) AND NOT xStop,
    diConnectID := cdiConnectID, pSend := pSend, uiSendSize := uiSendSize);
fbClose(xExecute := (uiStep = UINT#90) AND xOwned, diConnectID := cdiConnectID);
fbReplyTime(IN := (uiStep = UINT#30) OR (uiStep = UINT#40), PT := T#1s);
fbCloseTime(IN := (uiStep = UINT#90) AND xOwned, PT := T#3s);
fbPollTime(IN := uiStep = UINT#50, PT := T#100ms);
fbRetryTime(IN := uiStep = UINT#100, PT := T#1s);
CASE uiStep OF
    UINT#0:
        IF xEnable AND (uiPort > UINT#0) AND (byUnit > BYTE#0) AND (byUnit <= BYTE#247) THEN
            sRunAddress := sAddress; uiRunPort := uiPort; byRunUnit := byUnit;
            stServer.strIPAddr := sRunAddress; stServer.uiPort := uiRunPort;
            xError := FALSE; wErrorID := WORD#0;
            uiStep := UINT#10;
        END_IF;
    UINT#10:
        // Do not cancel a pending native connect before its terminal result.
        IF fbClient.xError THEN
            xError := TRUE; wErrorID := fbClient.wErrorID; uiStep := UINT#100;
        ELSIF fbClient.xDone THEN
            xOwned := TRUE;
            IF xStop THEN uiStep := UINT#90; ELSE uiStep := UINT#20; END_IF;
        END_IF;
    UINT#20:
        IF uiTransaction = UINT#65535 THEN uiTransaction := UINT#1;
        ELSE uiTransaction := uiTransaction + UINT#1; END_IF;
        aRequest[0] := UINT_TO_BYTE(SHR(uiTransaction,8));
        aRequest[1] := UINT_TO_BYTE(uiTransaction AND UINT#255);
        aRequest[2] := BYTE#0; aRequest[3] := BYTE#0;
        aRequest[4] := BYTE#0; aRequest[5] := BYTE#6;
        aRequest[6] := byRunUnit; aRequest[7] := BYTE#4;
        aRequest[8] := BYTE#0; aRequest[9] := BYTE#64;
        aRequest[10] := BYTE#0; aRequest[11] := BYTE#12;
        uiSent := UINT#0; uiReceived := UINT#0; uiStep := UINT#30;
    UINT#30:
        IF fbIo.xError OR fbIo.xPeerClosed OR fbReplyTime.Q THEN
            xFail := TRUE; wErrorID := WORD#16#A101;
        ELSE
            uiSent := uiSent + fbIo.uiSent;
            IF uiSent = UINT#12 THEN uiStep := UINT#40; END_IF;
        END_IF;
    UINT#40:
        IF fbIo.xError OR fbIo.xPeerClosed OR fbReplyTime.Q THEN
            xFail := TRUE; wErrorID := WORD#16#A102;
        ELSIF fbIo.uiCount > UINT#0 THEN
            IF uiReceived + fbIo.uiCount > UINT#33 THEN
                xFail := TRUE; wErrorID := WORD#16#A103;
            ELSE
                FOR i := UINT#0 TO fbIo.uiCount - UINT#1 DO
                    aResponse[uiReceived + i] := fbIo.aRecv[i];
                END_FOR;
                uiReceived := uiReceived + fbIo.uiCount;
                // Fail promptly on an exception or a malformed MBAP header.
                IF uiReceived >= UINT#9 THEN
                    IF (aResponse[0] <> aRequest[0]) OR (aResponse[1] <> aRequest[1])
                        OR (aResponse[2] <> BYTE#0) OR (aResponse[3] <> BYTE#0)
                        OR (aResponse[4] <> BYTE#0) OR (aResponse[5] <> BYTE#27)
                        OR (aResponse[6] <> byRunUnit) OR (aResponse[7] <> BYTE#4)
                        OR (aResponse[8] <> BYTE#24) THEN
                        xFail := TRUE; wErrorID := WORD#16#A104;
                    ELSIF uiReceived = UINT#33 THEN
                        FOR i := UINT#0 TO UINT#11 DO
                            aWords[i] := SHL(BYTE_TO_WORD(aResponse[9 + i*UINT#2]),8)
                                OR BYTE_TO_WORD(aResponse[10 + i*UINT#2]);
                        END_FOR;
                        IF udiCounter = UDINT#4294967295 THEN udiCounter := UDINT#1;
                        ELSE udiCounter := udiCounter + UDINT#1; END_IF;
                        xValid := TRUE; xUpdated := TRUE; xError := FALSE;
                        wErrorID := WORD#0; uiStep := UINT#50;
                    END_IF;
                END_IF;
            END_IF;
        END_IF;
    UINT#50:
        IF fbPollTime.Q THEN uiStep := UINT#20; END_IF;
    UINT#90:
        IF NOT xOwned THEN uiStep := UINT#100;
        ELSIF fbClose.xError OR fbCloseTime.Q THEN
            xCleanupFault := TRUE; xError := TRUE;
            wErrorID := WORD#16#A105; uiStep := UINT#200;
        ELSIF fbClose.xDone THEN xOwned := FALSE; uiStep := UINT#100; END_IF;
    UINT#100:
        IF fbRetryTime.Q THEN uiStep := UINT#0; END_IF;
    UINT#200:
        // A failed close keeps ownership latched. Never reuse or leak socket244.
        xValid := FALSE;
END_CASE;
IF xFail THEN xValid := FALSE; xError := TRUE; uiStep := UINT#90; END_IF;
IF xStop AND (uiStep <> UINT#0) AND (uiStep <> UINT#10)
    AND (uiStep <> UINT#90) AND (uiStep <> UINT#100) AND (uiStep <> UINT#200) THEN
    xValid := FALSE; uiStep := UINT#90;
END_IF;
fbAge(IN := NOT xUpdated, PT := T#1500ms);
uiAgeMs := UDINT_TO_UINT(TIME_TO_UDINT(fbAge.ET));
IF fbAge.Q OR NOT xEnable THEN xValid := FALSE; END_IF;
END_FUNCTION_BLOCK

(* ---- PRG_FileBridge.st ---- *)
PROGRAM PRG_FileBridge
VAR
    xInit : BOOL;
    xResetOld : BOOL;
    aPrevious : ARRAY[0..119] OF WORD;
    aSeen : ARRAY[0..119] OF WORD;
    aFrame : ARRAY[0..119] OF WORD;
    aAccepted : ARRAY[0..119] OF WORD;
    aFrameBytes : ARRAY[0..235] OF BYTE;
    aPayload : ARRAY[0..191] OF BYTE;
    aNames : ARRAY[0..31] OF STRING(64);
    uiState : UINT;
    wError : WORD;
    udiOwner : UDINT;
    udiAck : UDINT;
    uiAckOp : UINT;
    udiSize : UDINT;
    udiReceived : UDINT;
    udiExpectedCrc : UDINT;
    udiRunningCrc : UDINT := UDINT#16#FFFFFFFF;
    udiTotalSize : UDINT;
    uiVerified : UINT;
    uiExpectedFiles : UINT;
    uiOrdinal : UINT;
    uiMode : UINT;
    sProject : STRING(64);
    sFile : STRING(64);
    fbFtp : FB_FileFtp;
    fbLease : TON;
    wHeartbeatOld : WORD;
    xKick : BOOL;
    xStable : BOOL;
    xNew : BOOL;
    xSame : BOOL;
    xAccept : BOOL;
    xActive : BOOL;
    xClean : BOOL;
    xFileVerified : BOOL;
    xFtpStarted : BOOL;
    wReject : WORD;
    udiRejectSeq : UDINT;
    udiRejectOwner : UDINT;
    wRequestError : WORD;
    udiSeq : UDINT;
    udiSession : UDINT;
    udiBoot : UDINT;
    udiFrameCrc : UDINT;
    udiFrameSize : UDINT;
    udiOffset : UDINT;
    udiFileCrc : UDINT;
    uiOp : UINT;
    uiLength : UINT;
    uiCount : UINT;
    uiIndex : UINT;
    uiField : UINT;
    uiPos : UINT;
    uiI : UINT;
    uiJ : UINT;
    uiSnapshot : UINT;
    wFlags : WORD;
    sNewProject : STRING(64);
    sNewFile : STRING(64);
    pName : POINTER TO BYTE;
    xNamesOk : BOOL;
    xPairsOk : BOOL;
    xFound : BOOL;
    xGlobal : BOOL;
    uiPrograms : UINT;
    sPair : STRING(64);
    sReadyProject : STRING(64);
    uiReadyCapture : UINT;
    uiReadyPath : UINT;
    uiReadyReturn : UINT;
    xFixedConfig : BOOL;
    udiFixedProjectCrc : UDINT;
    uiSessionCapture : UINT;
    uiSessionPath : UINT;
    uiSessionReturn : UINT;
    aSessionTag : ARRAY[0..2] OF WORD;
END_VAR

(* This program NEVER writes robot motion/control outputs or GDI selection. *)
IF NOT xInit THEN
    GVL_FileBridge.xFixedReady := FALSE;
    GVL_FileBridge.xFixedUpdateBusy := FALSE;
    IF GVL_FileBridgeRetain.udiBootCounter = UDINT#16#FFFFFFFF THEN
        GVL_FileBridgeRetain.udiBootCounter := UDINT#1;
    ELSE
        GVL_FileBridgeRetain.udiBootCounter := GVL_FileBridgeRetain.udiBootCounter + UDINT#1;
    END_IF;
    FOR uiI := UINT#0 TO UINT#119 DO
        aPrevious[uiI] := GVL_FileBridge.aCommand[uiI];
        aSeen[uiI] := GVL_FileBridge.aCommand[uiI];
    END_FOR;
    xInit := TRUE;
END_IF;

xFixedConfig := GVL_FileBridge.xFixedMappingConfirmed
    AND (GVL_RobotBridge.uiFixedJobGuardVersion = UINT#140)
    AND F_FileNameValid(GVL_FileBridge.sFixedProject, TRUE)
    AND (GVL_FileBridge.uiFixedCapture >= UINT#1) AND (GVL_FileBridge.uiFixedCapture <= UINT#255)
    AND (GVL_FileBridge.uiFixedPath >= UINT#1) AND (GVL_FileBridge.uiFixedPath <= UINT#255)
    AND (GVL_FileBridge.uiAutoCapacity = UINT#15)
    AND (GVL_FileBridge.uiFixedCapture = UINT#10)
    AND (GVL_FileBridge.uiFixedPath <> UINT#10)
    AND (GVL_FileBridge.uiFixedCapture <> GVL_FileBridge.uiFixedPath)
;
GVL_FileBridge.xFixedIdle := GVL_RobotBridge.xRobotLinkOK AND GVL_RobotBridge.xRobotStopped
    AND NOT GVL_RobotBridge.xRobotRunning AND NOT GVL_RobotBridge.xRobotPaused
    AND NOT GVL_RobotBridge.xRobotEnabled AND NOT GVL_RobotBridge.xBusy
    AND NOT GVL_ManualBridge.xActive;
IF NOT xFixedConfig OR (sReadyProject <> GVL_FileBridge.sFixedProject)
    OR (uiReadyCapture <> GVL_FileBridge.uiFixedCapture) OR (uiReadyPath <> GVL_FileBridge.uiFixedPath)
    OR (uiReadyReturn <> GVL_FileBridge.uiAutoCapacity) THEN
    GVL_FileBridge.xFixedReady := FALSE;
END_IF;
udiFixedProjectCrc := F_FileCrc32(ADR(GVL_FileBridge.sFixedProject),
    INT_TO_UINT(LEN(GVL_FileBridge.sFixedProject)), UDINT#16#FFFFFFFF) XOR UDINT#16#FFFFFFFF;

xClean := NOT fbFtp.xControlOwned AND NOT fbFtp.xDataOwned
    AND ((fbFtp.uiStep = UINT#0) OR (fbFtp.uiStep = UINT#100));
IF GVL_FileBridge.xReset AND NOT xResetOld AND xClean
    AND (uiState <> UINT#300) AND (uiState <> UINT#310) THEN
    uiState := UINT#0;
    wError := WORD#0;
    udiOwner := UDINT#0;
    udiAck := UDINT#0;
    uiAckOp := UINT#0;
    uiVerified := UINT#0;
    uiExpectedFiles := UINT#0;
    udiReceived := UDINT#0;
    udiSize := UDINT#0;
    xFileVerified := FALSE;
    GVL_FileBridge.xFixedReady := FALSE;
    wReject := WORD#0;
END_IF;
xResetOld := GVL_FileBridge.xReset;

xActive := (uiState = UINT#100) OR (uiState = UINT#200)
    OR (uiState = UINT#300) OR (uiState = UINT#310);
xKick := FALSE;
IF (GVL_FileBridge.aHeartbeat[0] = UDINT_TO_WORD(SHR(udiOwner, 16)))
    AND (GVL_FileBridge.aHeartbeat[1] = UDINT_TO_WORD(udiOwner))
    AND (GVL_FileBridge.aHeartbeat[2] = UDINT_TO_WORD(SHR(GVL_FileBridgeRetain.udiBootCounter, 16)))
    AND (GVL_FileBridge.aHeartbeat[3] = UDINT_TO_WORD(GVL_FileBridgeRetain.udiBootCounter))
    AND (GVL_FileBridge.aHeartbeat[4] <> wHeartbeatOld) THEN
    wHeartbeatOld := GVL_FileBridge.aHeartbeat[4];
    xKick := TRUE;
END_IF;
fbLease(IN := xActive AND NOT xKick, PT := T#10s);

(* Two consecutive identical samples, then CRC of big-endian WORD bytes. *)
xStable := TRUE;
xNew := FALSE;
FOR uiI := UINT#0 TO UINT#119 DO
    aFrame[uiI] := GVL_FileBridge.aCommand[uiI];
    IF aFrame[uiI] <> aPrevious[uiI] THEN xStable := FALSE; END_IF;
    IF aFrame[uiI] <> aSeen[uiI] THEN xNew := TRUE; END_IF;
    aPrevious[uiI] := aFrame[uiI];
END_FOR;
IF xStable AND xNew THEN
    FOR uiI := UINT#0 TO UINT#119 DO aSeen[uiI] := aFrame[uiI]; END_FOR;
    FOR uiI := UINT#0 TO UINT#117 DO
        aFrameBytes[uiI * UINT#2] := WORD_TO_BYTE(SHR(aFrame[uiI], 8));
        aFrameBytes[uiI * UINT#2 + UINT#1] := WORD_TO_BYTE(aFrame[uiI] AND WORD#255);
    END_FOR;
    FOR uiI := UINT#0 TO UINT#95 DO
        aPayload[uiI * UINT#2] := WORD_TO_BYTE(SHR(aFrame[uiI + UINT#20], 8));
        aPayload[uiI * UINT#2 + UINT#1] := WORD_TO_BYTE(aFrame[uiI + UINT#20] AND WORD#255);
    END_FOR;
    uiOp := WORD_TO_UINT(aFrame[2]);
    udiSeq := SHL(WORD_TO_UDINT(aFrame[3]), 16) OR WORD_TO_UDINT(aFrame[4]);
    udiSession := SHL(WORD_TO_UDINT(aFrame[5]), 16) OR WORD_TO_UDINT(aFrame[6]);
    udiBoot := SHL(WORD_TO_UDINT(aFrame[7]), 16) OR WORD_TO_UDINT(aFrame[8]);
    udiFrameSize := SHL(WORD_TO_UDINT(aFrame[9]), 16) OR WORD_TO_UDINT(aFrame[10]);
    udiOffset := SHL(WORD_TO_UDINT(aFrame[11]), 16) OR WORD_TO_UDINT(aFrame[12]);
    uiLength := WORD_TO_UINT(aFrame[13]);
    udiFileCrc := SHL(WORD_TO_UDINT(aFrame[14]), 16) OR WORD_TO_UDINT(aFrame[15]);
    udiFrameCrc := F_FileCrc32(ADR(aFrameBytes), UINT#236, UDINT#16#FFFFFFFF) XOR UDINT#16#FFFFFFFF;
    wRequestError := WORD#0;
    xAccept := FALSE;
    IF (aFrame[0] <> WORD#16#F7B1) OR (aFrame[1] <> WORD#1)
        OR (((uiOp <> UINT#1) OR ((aFrame[18] <> WORD#2) AND (aFrame[18] <> WORD#3)))
            AND ((aFrame[19] <> WORD#0) OR (aFrame[116] <> WORD#0) OR (aFrame[117] <> WORD#0)))
        OR (uiLength > UINT#192) OR (udiSeq = UDINT#0) OR (udiSession = UDINT#0) THEN
        wRequestError := WORD#16#E001;
    ELSIF udiFrameCrc <> (SHL(WORD_TO_UDINT(aFrame[118]), 16) OR WORD_TO_UDINT(aFrame[119])) THEN
        wRequestError := WORD#16#E002;
    ELSIF udiBoot <> GVL_FileBridgeRetain.udiBootCounter THEN
        wRequestError := WORD#16#E003;
    ELSIF (udiSession = udiOwner) AND (udiSeq = udiAck) THEN
        xSame := TRUE;
        FOR uiI := UINT#0 TO UINT#119 DO
            IF aAccepted[uiI] <> aFrame[uiI] THEN xSame := FALSE; END_IF;
        END_FOR;
        IF NOT xSame THEN wRequestError := WORD#16#E004; END_IF;
        (* Exact replay: existing ACK/status only; NEVER repeat file/FTP operations. *)
    ELSE
        IF (uiOp = UINT#1) AND ((uiState = UINT#0) OR (uiState = UINT#400)) THEN
            IF (udiSeq <> UDINT#1) OR NOT xClean THEN wRequestError := WORD#16#E005; END_IF;
        ELSIF udiSession <> udiOwner THEN
            wRequestError := WORD#16#E006;
        ELSIF (udiSeq <= udiAck) OR (udiAck = UDINT#16#FFFFFFFF) THEN
            wRequestError := WORD#16#E005;
        ELSIF (uiOp <> UINT#4) AND (uiOp <> UINT#6) AND (udiSeq <> udiAck + UDINT#1) THEN
            wRequestError := WORD#16#E005;
        END_IF;
        IF NOT GVL_FileBridge.xFileTransferPermit AND (uiOp <> UINT#4) AND (uiOp <> UINT#6) THEN
            wRequestError := WORD#16#E007;
        END_IF;
        IF wRequestError = WORD#0 THEN
            CASE uiOp OF
                UINT#1: (* START file; first file also creates project session. *)
                    sNewProject := '';
                    sNewFile := '';
                    uiField := UINT#0;
                    uiPos := UINT#0;
                    xNamesOk := (uiLength >= UINT#2) AND (uiLength <= UINT#98);
                    IF xNamesOk THEN
                        FOR uiI := UINT#0 TO uiLength - UINT#1 DO
                            IF uiField = UINT#0 THEN pName := ADR(sNewProject);
                            ELSE pName := ADR(sNewFile); END_IF;
                            IF aPayload[uiI] = BYTE#0 THEN
                                IF uiPos = UINT#0 THEN xNamesOk := FALSE; END_IF;
                                uiField := uiField + UINT#1;
                                uiPos := UINT#0;
                            ELSIF (uiField > UINT#1) OR (uiPos >= UINT#48) THEN
                                xNamesOk := FALSE;
                            ELSE
                                pName[uiPos] := aPayload[uiI];
                                uiPos := uiPos + UINT#1;
                                pName[uiPos] := BYTE#0;
                            END_IF;
                        END_FOR;
                    END_IF;
                    xNamesOk := xNamesOk AND (uiField = UINT#2) AND (uiPos = UINT#0)
                        AND F_FileNameValid(sNewProject, TRUE) AND F_FileNameValid(sNewFile, FALSE);
                    uiCount := WORD_TO_UINT(aFrame[16]);
                    uiIndex := WORD_TO_UINT(aFrame[17]);
                    IF NOT GVL_FileBridge.xFileTransferPermit THEN
                        wRequestError := WORD#16#E007;
                    ELSIF NOT xNamesOk OR (aFrame[18] > WORD#3) THEN
                        wRequestError := WORD#16#E008;
                    ELSIF ((aFrame[18] = WORD#2) OR (aFrame[18] = WORD#3)) AND (NOT xFixedConfig
                        OR NOT GVL_FileBridge.xFixedIdle OR (sNewProject <> GVL_FileBridge.sFixedProject)
                        OR (uiCount < UINT#4) OR (uiCount > UINT#32) OR ((uiCount MOD UINT#2) <> UINT#0)
                        OR NOT F_FixedFileValid(sNewFile)
                        OR (aFrame[19] = WORD#0) OR (aFrame[19] > WORD#32767)
                        OR (aFrame[116] = WORD#0) OR (aFrame[116] > WORD#32767)
                        OR (aFrame[117] = WORD#0) OR (aFrame[117] > WORD#32767)) THEN
                        wRequestError := WORD#16#E015;
                    ELSIF ((aFrame[18] <> WORD#2) AND (aFrame[18] <> WORD#3)) AND (sNewProject = GVL_FileBridge.sFixedProject) THEN
                        wRequestError := WORD#16#E015;
                    ELSIF (udiFrameSize > UDINT#1048576)
                        OR (uiCount = UINT#0) OR (uiCount > UINT#32) OR (udiOffset <> UDINT#0) THEN
                        wRequestError := WORD#16#E009;
                    ELSIF (aFrame[18] = WORD#1) AND (RIGHT(sNewFile, 4) = '.txt') THEN
                        wRequestError := WORD#16#E008;
                    ELSIF (uiState = UINT#0) OR (uiState = UINT#400) THEN
                        IF (uiIndex <> UINT#1) OR (udiSeq <> UDINT#1) THEN
                            wRequestError := WORD#16#E00A;
                        ELSE
                            udiOwner := udiSession;
                            uiVerified := UINT#0;
                            udiTotalSize := UDINT#0;
                            uiExpectedFiles := uiCount;
                            uiMode := WORD_TO_UINT(aFrame[18]);
                            sProject := sNewProject;
                            IF uiMode >= UINT#2 THEN
                                GVL_FileBridge.xFixedReady := FALSE;
                                GVL_FileBridge.xFixedUpdateBusy := TRUE;
                                uiSessionCapture := GVL_FileBridge.uiFixedCapture;
                                uiSessionPath := GVL_FileBridge.uiFixedPath;
                                uiSessionReturn := GVL_FileBridge.uiAutoCapacity;
                                aSessionTag[0] := aFrame[19]; aSessionTag[1] := aFrame[116]; aSessionTag[2] := aFrame[117];
                            END_IF;
                            xAccept := TRUE;
                        END_IF;
                    ELSIF (uiState <> UINT#200) OR (sNewProject <> sProject)
                        OR (uiIndex <> uiVerified + UINT#1) OR (uiIndex > uiExpectedFiles)
                        OR (uiCount <> uiExpectedFiles) OR (aFrame[18] <> UINT_TO_WORD(uiMode)) THEN
                        wRequestError := WORD#16#E00A;
                    ELSE
                        xAccept := TRUE;
                        IF (uiMode >= UINT#2) AND ((aSessionTag[0] <> aFrame[19])
                            OR (aSessionTag[1] <> aFrame[116]) OR (aSessionTag[2] <> aFrame[117])) THEN
                            xAccept := FALSE; wRequestError := WORD#16#E015;
                        END_IF;
                        FOR uiI := UINT#0 TO uiVerified - UINT#1 DO
                            IF aNames[uiI] = sNewFile THEN
                                xAccept := FALSE;
                                wRequestError := WORD#16#E00B;
                            END_IF;
                        END_FOR;
                    END_IF;
                    IF xAccept THEN
                        IF udiTotalSize + udiFrameSize > UDINT#5242880 THEN
                            xAccept := FALSE;
                            wRequestError := WORD#16#E009;
                        ELSE
                            sFile := sNewFile;
                            udiSize := udiFrameSize;
                            udiExpectedCrc := udiFileCrc;
                            udiRunningCrc := UDINT#16#FFFFFFFF;
                            udiReceived := UDINT#0;
                            uiOrdinal := uiIndex;
                            uiState := UINT#100;
                            wError := WORD#0;
                            xFileVerified := FALSE;
                        END_IF;
                    END_IF;
                UINT#2: (* CHUNK; sequential, no writes while FTP owns buffer. *)
                    IF (uiMode = UINT#3) OR (uiState <> UINT#100) OR (uiLength = UINT#0)
                        OR (udiOffset <> udiReceived) OR (udiOffset + UINT_TO_UDINT(uiLength) > udiSize) THEN
                        wRequestError := WORD#16#E00C;
                    ELSE
                        FOR uiI := UINT#0 TO uiLength - UINT#1 DO
                            GVL_FileBridge.aBuffer[udiReceived + UINT_TO_UDINT(uiI)] := aPayload[uiI];
                        END_FOR;
                        udiRunningCrc := F_FileCrc32(ADR(aPayload), uiLength, udiRunningCrc);
                        udiReceived := udiReceived + UINT_TO_UDINT(uiLength);
                        xAccept := TRUE;
                    END_IF;
                UINT#3: (* DEPLOY only complete, CRC-checked RAM image. *)
                    IF (uiState <> UINT#100) OR ((uiMode <> UINT#3) AND (udiReceived <> udiSize)) OR (uiLength <> UINT#0) THEN
                        wRequestError := WORD#16#E00D;
                    ELSIF (uiMode <> UINT#3) AND ((udiRunningCrc XOR UDINT#16#FFFFFFFF) <> udiExpectedCrc) THEN
                        wRequestError := WORD#16#E00E;
                        wError := wRequestError;
                        uiState := UINT#900;
                    ELSIF NOT GVL_FileBridge.xFileTransferPermit THEN
                        wRequestError := WORD#16#E007;
                    ELSE
                        uiState := UINT#300;
                        xAccept := TRUE;
                    END_IF;
                UINT#4: (* ABORT; cleanup cannot be skipped or rearmed remotely. *)
                    IF (uiState = UINT#300) OR (uiState = UINT#310) THEN
                        uiState := UINT#310;
                    ELSE
                        uiState := UINT#900;
                    END_IF;
                    wError := WORD#16#E010;
                    xAccept := TRUE;
                UINT#5: (* FINISH: all files individually uploaded AND read back. *)
                    IF (uiState <> UINT#200) OR (uiVerified <> uiExpectedFiles) THEN
                        wRequestError := WORD#16#E00F;
                    ELSIF (uiMode >= UINT#2) AND (NOT xFixedConfig OR NOT GVL_FileBridge.xFixedIdle
                        OR (sProject <> GVL_FileBridge.sFixedProject)
                        OR (uiSessionCapture <> GVL_FileBridge.uiFixedCapture)
                        OR (uiSessionPath <> GVL_FileBridge.uiFixedPath)
                        OR (uiSessionReturn <> GVL_FileBridge.uiAutoCapacity)) THEN
                        wRequestError := WORD#16#E015;
                    ELSE
                        xPairsOk := TRUE;
                        IF uiMode = UINT#1 THEN
                            xGlobal := FALSE;
                            uiPrograms := UINT#0;
                            FOR uiI := UINT#0 TO uiVerified - UINT#1 DO
                                IF aNames[uiI] = '_project.srd' THEN xGlobal := TRUE; END_IF;
                                IF RIGHT(aNames[uiI], 4) = '.srp' THEN
                                    uiPrograms := uiPrograms + UINT#1;
                                    sPair := CONCAT(LEFT(aNames[uiI], LEN(aNames[uiI]) - 1), 'd');
                                    xFound := FALSE;
                                    FOR uiJ := UINT#0 TO uiVerified - UINT#1 DO
                                        IF aNames[uiJ] = sPair THEN xFound := TRUE; END_IF;
                                    END_FOR;
                                    IF NOT xFound THEN xPairsOk := FALSE; END_IF;
                                END_IF;
                            END_FOR;
                            xPairsOk := xPairsOk AND xGlobal AND (uiPrograms > UINT#0);
                        END_IF;
                        IF uiMode >= UINT#2 THEN
                            FOR uiI := UINT#0 TO uiVerified - UINT#1 DO
                                IF (F_AutoFileIndex(aNames[uiI]) = UINT#0)
                                    OR (F_AutoFileIndex(aNames[uiI]) > uiVerified) THEN xPairsOk := FALSE; END_IF;
                            END_FOR;
                        END_IF;
                        IF xPairsOk THEN
                            uiState := UINT#400; xAccept := TRUE;
                            IF uiMode >= UINT#2 THEN
                                GVL_FileBridge.xFixedReady := TRUE;
                                FOR uiI := UINT#0 TO UINT#2 DO GVL_FileBridge.aAutoTag[uiI] := aSessionTag[uiI]; END_FOR;
                                sReadyProject := GVL_FileBridge.sFixedProject;
                                uiReadyCapture := GVL_FileBridge.uiFixedCapture;
                                uiReadyPath := GVL_FileBridge.uiFixedPath;
                                uiReadyReturn := GVL_FileBridge.uiAutoCapacity;
                            END_IF;
                        ELSE wRequestError := WORD#16#E012; END_IF;
                    END_IF;
                UINT#6: (* RELEASE only after all handles are known closed. *)
                    IF xClean AND ((uiState = UINT#400) OR (uiState = UINT#900)) THEN
                        uiState := UINT#0;
                        xAccept := TRUE;
                    ELSE wRequestError := WORD#16#E013; END_IF;
            ELSE
                wRequestError := WORD#16#E001;
            END_CASE;
        END_IF;
        IF xAccept THEN
            udiAck := udiSeq;
            uiAckOp := uiOp;
            FOR uiI := UINT#0 TO UINT#119 DO aAccepted[uiI] := aFrame[uiI]; END_FOR;
        END_IF;
    END_IF;
    IF wRequestError <> WORD#0 THEN
        wReject := wRequestError;
        udiRejectSeq := udiSeq;
        udiRejectOwner := udiSession;
    END_IF;
END_IF;

IF xActive AND (fbLease.Q OR NOT GVL_FileBridge.xFileTransferPermit
    OR ((uiMode >= UINT#2) AND (NOT xFixedConfig OR NOT GVL_FileBridge.xFixedIdle
        OR (sProject <> GVL_FileBridge.sFixedProject)
        OR (uiSessionCapture <> GVL_FileBridge.uiFixedCapture)
        OR (uiSessionPath <> GVL_FileBridge.uiFixedPath)
        OR (uiSessionReturn <> GVL_FileBridge.uiAutoCapacity)))) THEN
    IF fbLease.Q THEN wError := WORD#16#E011;
    ELSE wError := WORD#16#E007; END_IF;
    IF (uiState = UINT#300) OR (uiState = UINT#310) THEN uiState := UINT#310;
    ELSIF uiState <> UINT#400 THEN uiState := UINT#900; END_IF;
END_IF;

IF ((uiState = UINT#300) OR (uiState = UINT#310)) AND xFtpStarted AND fbFtp.xDone THEN
    xFtpStarted := FALSE;
    IF (uiState = UINT#300) AND fbFtp.xTestPassed THEN
        IF uiMode = UINT#3 THEN
            (* FB CRC was verified against this session's immutable expected CRC. *)
            udiRunningCrc := udiExpectedCrc XOR UDINT#16#FFFFFFFF;
        END_IF;
        aNames[uiVerified] := sFile;
        uiVerified := uiVerified + UINT#1;
        udiTotalSize := udiTotalSize + udiSize;
        xFileVerified := TRUE;
        uiState := UINT#200;
    ELSE
        IF wError = WORD#0 THEN wError := WORD#16#E014; END_IF;
        IF fbFtp.xControlOwned OR fbFtp.xDataOwned THEN uiState := UINT#910;
        ELSE uiState := UINT#900; END_IF;
    END_IF;
END_IF;
IF (uiState = UINT#300) OR (uiState = UINT#310) THEN xFtpStarted := TRUE; END_IF;
fbFtp(xStart := (uiState = UINT#300) OR (uiState = UINT#310),
    xAbort := uiState = UINT#310, pBuffer := ADR(GVL_FileBridge.aBuffer),
    udiSize := udiSize, sProject := sProject, sFile := sFile,
    xCreateProject := uiVerified = UINT#0,
    xReplaceFixed := uiMode >= UINT#2,
    xVerifyOnly := uiMode = UINT#3, udiVerifyCrc := udiExpectedCrc,
    sUser := GVL_FileBridge.sFtpUser, sPassword := GVL_FileBridge.sFtpPassword);

(* Coherent FC03 status: matching EVEN snapshot head/tail required by PC. *)
IF uiSnapshot >= UINT#65534 THEN uiSnapshot := UINT#0;
ELSE uiSnapshot := uiSnapshot + UINT#2; END_IF;
GVL_FileBridge.aStatus[38] := UINT_TO_WORD(uiSnapshot + UINT#1);
wFlags := WORD#0;
IF GVL_FileBridge.xFileTransferPermit THEN wFlags := wFlags OR WORD#1; END_IF;
IF xClean THEN wFlags := wFlags OR WORD#2; END_IF;
IF xFileVerified THEN wFlags := wFlags OR WORD#4; END_IF;
IF uiState = UINT#400 THEN wFlags := wFlags OR WORD#8; END_IF;
IF (uiState = UINT#300) OR (uiState = UINT#310) THEN wFlags := wFlags OR WORD#16; END_IF;
GVL_FileBridge.aStatus[0] := WORD#16#F7B2;
GVL_FileBridge.aStatus[1] := WORD#1;
GVL_FileBridge.aStatus[2] := UINT_TO_WORD(uiState);
GVL_FileBridge.aStatus[3] := wError;
GVL_FileBridge.aStatus[4] := UDINT_TO_WORD(SHR(udiAck, 16));
GVL_FileBridge.aStatus[5] := UDINT_TO_WORD(udiAck);
GVL_FileBridge.aStatus[6] := UINT_TO_WORD(uiAckOp);
GVL_FileBridge.aStatus[7] := wFlags;
GVL_FileBridge.aStatus[8] := UDINT_TO_WORD(SHR(udiOwner, 16));
GVL_FileBridge.aStatus[9] := UDINT_TO_WORD(udiOwner);
GVL_FileBridge.aStatus[10] := UDINT_TO_WORD(SHR(GVL_FileBridgeRetain.udiBootCounter, 16));
GVL_FileBridge.aStatus[11] := UDINT_TO_WORD(GVL_FileBridgeRetain.udiBootCounter);
GVL_FileBridge.aStatus[12] := UDINT_TO_WORD(SHR(udiReceived, 16));
GVL_FileBridge.aStatus[13] := UDINT_TO_WORD(udiReceived);
GVL_FileBridge.aStatus[14] := UDINT_TO_WORD(SHR(udiSize, 16));
GVL_FileBridge.aStatus[15] := UDINT_TO_WORD(udiSize);
GVL_FileBridge.aStatus[16] := UDINT_TO_WORD(SHR(udiRunningCrc XOR UDINT#16#FFFFFFFF, 16));
GVL_FileBridge.aStatus[17] := UDINT_TO_WORD(udiRunningCrc XOR UDINT#16#FFFFFFFF);
GVL_FileBridge.aStatus[18] := UDINT_TO_WORD(SHR(udiExpectedCrc, 16));
GVL_FileBridge.aStatus[19] := UDINT_TO_WORD(udiExpectedCrc);
GVL_FileBridge.aStatus[20] := UINT_TO_WORD(uiVerified);
GVL_FileBridge.aStatus[21] := UINT_TO_WORD(uiExpectedFiles);
GVL_FileBridge.aStatus[22] := UINT_TO_WORD(uiOrdinal);
GVL_FileBridge.aStatus[23] := UINT_TO_WORD(fbFtp.uiStep);
GVL_FileBridge.aStatus[24] := UINT_TO_WORD(fbFtp.uiReplyCode);
GVL_FileBridge.aStatus[25] := fbFtp.wErrorID;
GVL_FileBridge.aStatus[26] := UINT_TO_WORD(fbFtp.uiErrorStage);
GVL_FileBridge.aStatus[27] := UDINT_TO_WORD(SHR(fbFtp.udiUploadedBytes, 16));
GVL_FileBridge.aStatus[28] := UDINT_TO_WORD(fbFtp.udiUploadedBytes);
GVL_FileBridge.aStatus[29] := UDINT_TO_WORD(SHR(fbFtp.udiReadbackBytes, 16));
GVL_FileBridge.aStatus[30] := UDINT_TO_WORD(fbFtp.udiReadbackBytes);
GVL_FileBridge.aStatus[31] := wReject;
GVL_FileBridge.aStatus[32] := UDINT_TO_WORD(SHR(udiRejectSeq, 16));
GVL_FileBridge.aStatus[33] := UDINT_TO_WORD(udiRejectSeq);
GVL_FileBridge.aStatus[34] := UDINT_TO_WORD(SHR(udiRejectOwner, 16));
GVL_FileBridge.aStatus[35] := UDINT_TO_WORD(udiRejectOwner);
GVL_FileBridge.aStatus[36] := wHeartbeatOld;
GVL_FileBridge.aStatus[37] := WORD#32;
GVL_FileBridge.aStatus[39] := WORD#16;
GVL_FileBridge.aStatus[40] := WORD#0;
GVL_FileBridge.aStatus[41] := WORD#192;
GVL_FileBridge.aStatus[42] := fbFtp.wDataCloseErrorID;
GVL_FileBridge.aStatus[43] := fbFtp.wControlCloseErrorID;
GVL_FileBridge.aStatus[44] := UINT_TO_WORD(uiMode);
GVL_FileBridge.aStatus[45] := UINT_TO_WORD(fbFtp.uiUploadCompleteCode);
GVL_FileBridge.aStatus[46] := UINT_TO_WORD(fbFtp.uiDownloadCompleteCode);
GVL_FileBridge.aStatus[47] := WORD#13; (* bit0 empty files; bit1 guarded fixed-project replacement *)
GVL_FileBridge.aStatus[48] := WORD#16#0104;
FOR uiI := UINT#49 TO UINT#62 DO GVL_FileBridge.aStatus[uiI] := WORD#0; END_FOR;
IF xFixedConfig THEN GVL_FileBridge.aStatus[49] := WORD#1; END_IF;
GVL_FileBridge.xFixedUpdateBusy := (uiMode >= UINT#2) AND ((uiState = UINT#100)
    OR (uiState = UINT#200) OR (uiState = UINT#300) OR (uiState = UINT#310) OR (uiState = UINT#910));
IF GVL_FileBridge.xFixedUpdateBusy THEN GVL_FileBridge.aStatus[50] := WORD#1; END_IF;
IF GVL_FileBridge.xFixedReady THEN GVL_FileBridge.aStatus[51] := WORD#1; END_IF;
GVL_FileBridge.aStatus[52] := UINT_TO_WORD(GVL_FileBridge.uiFixedCapture);
GVL_FileBridge.aStatus[53] := UINT_TO_WORD(GVL_FileBridge.uiFixedPath);
GVL_FileBridge.aStatus[54] := UINT_TO_WORD(GVL_FileBridge.uiAutoCapacity);
GVL_FileBridge.aStatus[55] := UDINT_TO_WORD(SHR(udiFixedProjectCrc, 16));
GVL_FileBridge.aStatus[56] := UDINT_TO_WORD(udiFixedProjectCrc);
IF GVL_FileBridge.xFixedIdle THEN GVL_FileBridge.aStatus[59] := WORD#1; END_IF;
GVL_FileBridge.aStatus[57] := GVL_FileBridge.aAutoTag[0];
GVL_FileBridge.aStatus[58] := GVL_FileBridge.aAutoTag[1];
GVL_FileBridge.aStatus[60] := GVL_FileBridge.aAutoTag[2];
GVL_FileBridge.aStatus[61] := WORD#8192;
GVL_FileBridge.aStatus[62] := WORD#1; (* batch I/O backend revision *)
(* Execute after ManualBridge: it clears the same parameter words first. *)
IF GVL_FileBridge.xFixedReady AND NOT GVL_ManualBridge.xActive
    AND (GVL_RobotBridge.aHostStatus[13] = UINT_TO_WORD(GVL_FileBridge.uiFixedPath)) THEN
    FOR uiI := UINT#0 TO UINT#2 DO GVL_ParamProbe.aParamTx[uiI] := GVL_FileBridge.aAutoTag[uiI]; END_FOR;
END_IF;
GVL_FileBridge.aStatus[63] := UINT_TO_WORD(uiSnapshot);
GVL_FileBridge.aStatus[38] := UINT_TO_WORD(uiSnapshot);
END_PROGRAM
